{attribute 'enable_dynamic_creation'}
FUNCTION_BLOCK FB_Dynamic
VAR
    nCounts : INT;
END_VAR

METHOD Increase : INT
VAR_INPUT
	nCountStep :INT;
END_VAR
nCounts := nCounts + nCountStep;
Increase := nCounts;
END_METHOD

END_FUNCTION_BLOCK

(* stored: Version 1.1.0.1, ProductVersion 3.1.4026.21
   POU FB_Dynamic: Id {1a9f2f1f-3aa5-4017-8184-8fb8a4cd4490}, SpecialFunc None
   Method Increase: Id {ef4ca4c5-48cb-4ca8-9490-f1291786189c} *)
